Fanuc KAREL source: KT00362.KL

PROGRAM KT00362
%NOLOCKGROUP
VAR
  P1: JOINTPOS
  P2: JOINTPOS
  OUT: BOOLEAN
BEGIN
  OUT = P1 < P2
END KT00362
